Fanuc KAREL source: kf00081.KL

-- PROVISIONAL review KL for V940-1; original PC SHA256 efb77a63c1717f2cf83a57077b2acd52d8778f3aa6db325c03923f010384ed3e
-- Incomplete behavior may be omitted. Consult companion uncertainty JSON. Do not deploy.
PROGRAM KF00081
%NOLOCKGROUP
BEGIN
  -- V9_ZERO_TABLE_METADATA_HINT layout=0002_ascii; no indexed target words; source/name/runtime held
  -- UNRESOLVED_PC offsets 5-15; opcodes 27,22,31
  -- UNRESOLVED_PC offsets 20-54; opcodes 27,27,2E,22,22,22,22,31
  -- UNRESOLVED_PC offsets 59-63; opcodes 7F
END KF00081
